// 	            (HMI_Box_Connected_2 = 34 AND KEY_REMOTE_LOCAL_L4___CH1_3_) OR
// 	            (HMI_Box_Connected_2 = 35 AND KEY_REMOTE_LOCAL_L5___CH1_3_) OR
// 	            (HMI_Box_Connected_2 = 36 AND KEY_REMOTE_LOCAL_L6___CH1_3_) OR
// 	            (HMI_Box_Connected_2 = 37 AND KEY_REMOTE_LOCAL_L7___CH1_3_) OR
// 	            (HMI_Box_Connected_2 = 38 AND KEY_REMOTE_LOCAL_L8___CH1_3_)
// 	        THEN
// 	            Errors_Profinet_3.%X8 :=
// 	            Errors_Profinet_5.%X0 :=
// 	            Errors_Profinet_5.%X2 :=
// 	            Errors_Profinet_5.%X3 :=
// 	            Errors_Profinet_5.%X4 :=
// 	            Errors_Profinet_5.%X5 :=
// 	            Errors_Profinet_5.%X6 :=
// 	            Errors_Profinet_5.%X7 :=
// 	            Errors_Profinet_5.%X8 :=
// 	            Errors_Profinet_5.%X9 :=
// 	            Errors_Profinet_5.%X10 :=
// 	            Errors_Profinet_5.%X12 :=
// 	            Errors_Profinet_5.%X13 :=
// 	            Errors_Profinet_5.%X14 :=
// 	            Errors_Profinet_5.%X15 :=
// 	            Errors_Profinet_6.%X0 :=
// 	            Errors_Profinet_6.%X1 :=
// 	            Errors_Profinet_6.%X2 :=
// 	            Errors_Profinet_6.%X3 :=
// 	            Errors_Profinet_6.%X4 :=
// 	            Errors_Profinet_6.%X5 :=
// 	            Errors_Profinet_6.%X6 :=
// 	            Errors_Profinet_6.%X7 :=
// 	            Errors_Profinet_6.%X8 :=
// 	            Errors_Profinet_6.%X9 :=
// 	            Errors_Profinet_6.%X10 :=
// 	            Errors_Profinet_6.%X11 :=
// 	            Errors_Profinet_7.%X2 :=
// 	            Errors_Profinet_8.%X7 :=
// 	            Errors_Profinet_9.%X7 :=
// 	            Errors_Profinet_9.%X8 :=
// 	            Errors_Profinet_9.%X9 :=
// 	            Errors_Profinet_9.%X10 :=
// 	            Errors_Profinet_10.%X2 :=
// 	            Errors_Profinet_10.%X3 :=
// 	            Errors_Profinet_10.%X4 :=
// 	            Errors_Profinet_10.%X5 :=
// 
// 	            Erros_Supply_Feedback_4.%X8 :=
// 	            Erros_Supply_Feedback_4.%X9 :=
// 	            Erros_Supply_Feedback_4.%X10 :=
// 	            Erros_Supply_Feedback_4.%X11 :=
// 	            Erros_Supply_Feedback_4.%X12 :=
// 	            Erros_Supply_Feedback_4.%X13 :=
// 	            Erros_Supply_Feedback_4.%X14 :=
// 	            Erros_Supply_Feedback_4.%X15 :=
// 	            Erros_Supply_Feedback_5.%X0 :=
// 	            Erros_Supply_Feedback_5.%X1 :=
// 	            Erros_Supply_Feedback_5.%X2 :=
// 	            Erros_Supply_Feedback_5.%X3 :=
// 	            Erros_Supply_Feedback_5.%X4 :=
// 	            Erros_Supply_Feedback_5.%X5 :=
// 	            Erros_Supply_Feedback_5.%X6 :=
// 	            Erros_Supply_Feedback_5.%X7 :=
// 	            Erros_Supply_Feedback_5.%X8 :=
// 	            Erros_Supply_Feedback_5.%X9 :=
// 	            Erros_Supply_Feedback_5.%X10 :=
// 	            Erros_Supply_Feedback_5.%X11 :=
// 
// 	            Estop_Error_Word_3.%X1 :=
// 	            Estop_Error_Word_3.%X2 :=
// 	            Estop_Error_Word_3.%X3 :=
// 	            Estop_Error_Word_3.%X4 :=
// 	            Estop_Error_Word_3.%X5 :=
// 	            Estop_Error_Word_3.%X6 :=
// 	            Estop_Error_Word_3.%X7 :=
// 	            Estop_Error_Word_3.%X8 :=
// 	            Estop_Error_Word_3.%X9 :=
// 	            Estop_Error_Word_3.%X10 :=
// 	            Estop_Error_Word_3.%X11 := FALSE;
// 
// 	            Sick_Lector_Error_code_3_2 :=
// 	            Linear_Encoder_Device_Errors_3 :=
// 	            Sick_Lector_Error_code_3 := 0;
// 
// 	            Errors_Word_LightGuard_1.%X4 := FALSE;
// 	            Errors_Word_LightGuard_1.%X5 := FALSE;
// 	        END_IF;
// 
// 
// 	        IF Screen_DB_1.Reset_All[2] AND
// 	            (HMI_Box_Connected_2 = 31 AND KEY_REMOTE_LOCAL_L1___CH1_3_) OR
// 	            (HMI_Box_Connected_2 = 32 AND KEY_REMOTE_LOCAL_L2___CH1_3_) OR
// 	            (HMI_Box_Connected_2 = 33 AND KEY_REMOTE_LOCAL_L3___CH1_3_) OR
// 	            (HMI_Box_Connected_2 = 34 AND KEY_REMOTE_LOCAL_L4___CH1_3_) OR
// 	            (HMI_Box_Connected_2 = 35 AND KEY_REMOTE_LOCAL_L5___CH1_3_) OR
// 	            (HMI_Box_Connected_2 = 36 AND KEY_REMOTE_LOCAL_L6___CH1_3_) OR
// 	            (HMI_Box_Connected_2 = 37 AND KEY_REMOTE_LOCAL_L7___CH1_3_) OR
// 	            (HMI_Box_Connected_2 = 38 AND KEY_REMOTE_LOCAL_L8___CH1_3_)
// 	        THEN
// 	            Errors_Profinet_3.%X8 :=
// 	            Errors_Profinet_5.%X5 :=
// 	            Errors_Profinet_6.%X13 :=
// 	            Errors_Profinet_6.%X15 :=
// 	            Errors_Profinet_7.%X0 :=
// 	            Errors_Profinet_7.%X1 :=
// 	            Errors_Profinet_7.%X2 :=
// 	            Errors_Profinet_7.%X3 :=
// 	            Errors_Profinet_7.%X4 :=
// 	            Errors_Profinet_7.%X5 :=
// 	            Errors_Profinet_7.%X6 :=
// 	            Errors_Profinet_7.%X7 :=
// 	            Errors_Profinet_7.%X8 :=
// 	            Errors_Profinet_7.%X9 :=
// 	            Errors_Profinet_7.%X10 :=
// 	            Errors_Profinet_7.%X11 :=
// 	            Errors_Profinet_7.%X12 :=
// 	            Errors_Profinet_7.%X13 :=
// 	            Errors_Profinet_7.%X14 :=
// 	            Errors_Profinet_7.%X15 :=
// 	            Errors_Profinet_8.%X0 :=
// 	            Errors_Profinet_8.%X7 :=
// 	            Errors_Profinet_9.%X7 :=
// 	            Errors_Profinet_9.%X8 :=
// 	            Errors_Profinet_9.%X9 :=
// 	            Errors_Profinet_9.%X10 :=
// 	            Errors_Profinet_10.%X6 :=
// 	            Errors_Profinet_10.%X7 :=
// 	            Errors_Profinet_10.%X8 :=
// 	            Errors_Profinet_10.%X9 :=
// 
// 	            Erros_Supply_Feedback_5.%X12 :=
// 	            Erros_Supply_Feedback_5.%X13 :=
// 	            Erros_Supply_Feedback_5.%X14 :=
// 	            Erros_Supply_Feedback_5.%X15 :=
// 	            Erros_Supply_Feedback_6.%X0 :=
// 	            Erros_Supply_Feedback_6.%X1 :=
// 	            Erros_Supply_Feedback_6.%X2 :=
// 	            Erros_Supply_Feedback_6.%X3 :=
// 	            Erros_Supply_Feedback_6.%X4 :=
// 	            Erros_Supply_Feedback_6.%X5 :=
// 	            Erros_Supply_Feedback_6.%X6 :=
// 	            Erros_Supply_Feedback_6.%X7 :=
// 
// 	            Estop_Error_Word_4.%X1 :=
// 	            Estop_Error_Word_4.%X2 :=
// 	            Estop_Error_Word_4.%X3 :=
// 	            Estop_Error_Word_4.%X4 :=
// 	            Estop_Error_Word_4.%X5 :=
// 	            Estop_Error_Word_4.%X6 :=
// 	            Estop_Error_Word_4.%X7 :=
// 	            Estop_Error_Word_4.%X8 :=
// 	            Estop_Error_Word_4.%X9 :=
// 	            Estop_Error_Word_4.%X10 := FALSE;
// 
// 	            Sick_Lector_Error_code_4_2 :=
// 	            Linear_Encoder_Device_Errors_4 :=
// 	            Sick_Lector_Error_code_4 := 0;
// 	        END_IF;
// 
// 
// 	        IF Screen_DB_1.Reset_All[2] AND
// 	            (HMI_Box_Connected_2 = 51 AND KEY_REMOTE_LOCAL_L1___CH1_5_) OR
// 	            (HMI_Box_Connected_2 = 52 AND KEY_REMOTE_LOCAL_L2___CH1_5_) OR
// 	            (HMI_Box_Connected_2 = 53 AND KEY_REMOTE_LOCAL_L3___CH1_5_) OR
// 	            (HMI_Box_Connected_2 = 54 AND KEY_REMOTE_LOCAL_L4___CH1_5_) OR
// 	            (HMI_Box_Connected_2 = 55 AND KEY_REMOTE_LOCAL_L5___CH1_5_) OR
// 	            (HMI_Box_Connected_2 = 56 AND KEY_REMOTE_LOCAL_L6___CH1_5_) OR
// 	            (HMI_Box_Connected_2 = 57 AND KEY_REMOTE_LOCAL_L7___CH1_5_) OR
// 	            (HMI_Box_Connected_2 = 58 AND KEY_REMOTE_LOCAL_L8___CH1_5_)
// 	        THEN
// 	            Errors_Profinet_3.%X8 :=
// 	            Errors_Profinet_5.%X5 :=
// 	            Errors_Profinet_7.%X2 :=
// 	            Errors_Profinet_8.%X2 :=
// 	            Errors_Profinet_8.%X4 :=
// 	            Errors_Profinet_8.%X5 :=
// 	            Errors_Profinet_8.%X6 :=
// 	            Errors_Profinet_8.%X7 :=
// 	            Errors_Profinet_8.%X8 :=
// 	            Errors_Profinet_8.%X9 :=
// 	            Errors_Profinet_8.%X10 :=
// 	            Errors_Profinet_8.%X11 :=
// 	            Errors_Profinet_8.%X12 :=
// 	            Errors_Profinet_8.%X13 :=
// 	            Errors_Profinet_8.%X14 :=
// 	            Errors_Profinet_8.%X15 :=
// 	            Errors_Profinet_9.%X0 :=
// 	            Errors_Profinet_9.%X1 :=
// 	            Errors_Profinet_9.%X2 :=
// 	            Errors_Profinet_9.%X3 :=
// 	            Errors_Profinet_9.%X4 :=
// 	            Errors_Profinet_9.%X5 :=
// 	            Errors_Profinet_9.%X7 :=
// 	            Errors_Profinet_9.%X8 :=
// 	            Errors_Profinet_9.%X9 :=
// 	            Errors_Profinet_9.%X10 :=
// 	            Errors_Profinet_10.%X10 :=
// 	            Errors_Profinet_10.%X11 :=
// 	            Errors_Profinet_10.%X12 :=
// 	            Errors_Profinet_10.%X13 :=
// 
// 	            Erros_Supply_Feedback_6.%X8 :=
// 	            Erros_Supply_Feedback_6.%X9 :=
// 	            Erros_Supply_Feedback_6.%X10 :=
// 	            Erros_Supply_Feedback_6.%X11 :=
// 	            Erros_Supply_Feedback_6.%X12 :=
// 	            Erros_Supply_Feedback_6.%X13 :=
// 	            Erros_Supply_Feedback_6.%X14 :=
// 	            Erros_Supply_Feedback_6.%X15 :=
// 	            Erros_Supply_Feedback_7.%X0 :=
// 	            Erros_Supply_Feedback_7.%X1 :=
// 	            Erros_Supply_Feedback_7.%X2 :=
// 	            Erros_Supply_Feedback_7.%X3 :=
// 
// 	            Estop_Error_Word_5.%X1 :=
// 	            Estop_Error_Word_5.%X2 :=
// 	            Estop_Error_Word_5.%X3 :=
// 	            Estop_Error_Word_5.%X4 :=
// 	            Estop_Error_Word_5.%X5 :=
// 	            Estop_Error_Word_5.%X6 :=
// 	            Estop_Error_Word_5.%X7 :=
// 	            Estop_Error_Word_5.%X8 :=
// 	            Estop_Error_Word_5.%X9 :=
// 	            Estop_Error_Word_5.%X10 := FALSE;
// 
// 	            Sick_Lector_Error_code_5_2 :=
// 	            Linear_Encoder_Device_Errors_5 :=
// 	            Sick_Lector_Error_code_5 := 0;
// 	        END_IF;

END_FUNCTION

(* stored: Version 1.1.0.1
   POU Errors_Warings: Id {d7669ad1-be00-5ba1-9310-bf776fe79181}, SpecialFunc None *)
